(* IEC 61131-3 sources: Repository_IEMA_Test/LMC_PacDrive.device.xml.v3^/Plc Logic.plclogic.xml.v3^/Application.application.xml.v3^/TemplateFullProgrammingFramework/Examples/ExampleLeafModule/FB_ExampleLeafModule.pou.xml.v3^, 16 files *)

(* ---- Auto_Action.act.st ---- *)
__METADATA__
{
  "v3Meta": {
    "objectGuid": "52a75849-8094-4c85-bfe0-08668a2e7324",
    "objectTypeGuid": "8ac092e5-3128-4e26-9e7e-11016c6684f2",
    "embeddedObjectTypeGuids": [
      "3b83b776-fb25-43b8-99f2-3c507c9143fc"
    ],
    "properties": {},
    "subObjects": {}
  }
}

(* Start application code *)
IF(iq_stExampleLeafModuleItf.q_etState = ET_ExampleLeafModuleState.AutoWaitForStart) THEN
	IF(xAutoEnable) THEN
		IF(xStartFlag) THEN
			iq_stExampleLeafModuleItf.q_etState := ET_ExampleLeafModuleState.AutoRunning;
		END_IF
	ELSE
		xAutoActive := FALSE;
	END_IF
END_IF

IF(NOT xStartFlag AND iq_stExampleLeafModuleItf.q_etState = ET_ExampleLeafModuleState.AutoRunning) THEN
	iq_stExampleLeafModuleItf.q_etState := ET_ExampleLeafModuleState.AutoWaitForStart;
END_IF

IF(iq_stExampleLeafModuleItf.q_etState = ET_ExampleLeafModuleState.AutoRunning) THEN
	IF(xAutoEnable) THEN
		iq_stExampleLeafModuleItf.q_xValue := ifRefActualValuesPosition.RefPosition >= iq_stExampleLeafModuleItf.i_lrPosMin AND
													ifRefActualValuesPosition.RefPosition <= iq_stExampleLeafModuleItf.i_lrPosMax;
	ELSE
		iq_stExampleLeafModuleItf.q_etState := ET_ExampleLeafModuleState.AutoWaitForStart;
	END_IF
END_IF
(* End application code *)

(* ---- CancelException.meth.st ---- *)
METHOD CancelException
VAR_IN_OUT
	iq_stException	: TPL.ST_Exception;
END_VAR

TPL.FC_SetException(	i_xExceptionActive	:= FALSE,
						iq_stException		:= iq_stException,
						iq_stExceptionList	:= iq_stExceptionList,
						iq_stLogDataList	:= iq_stLogDataList,
						q_etDiag 			=> etDiagBuffer,
						q_etDiagExt 		=> etDiagExtBufferTPL,
						q_sMsg 				=> sDiagMsgBuffer);

(* ---- CheckCmd.act.st ---- *)
__METADATA__
{
  "v3Meta": {
    "objectGuid": "c3140d7a-2c8d-489a-98e5-cdbf2202bc2d",
    "objectTypeGuid": "8ac092e5-3128-4e26-9e7e-11016c6684f2",
    "embeddedObjectTypeGuids": [
      "3b83b776-fb25-43b8-99f2-3c507c9143fc"
    ],
    "properties": {},
    "subObjects": {}
  }
}

(*--------------------------------------------------------------------------------------------------*)
(* CheckCMD is checking if CMD is supported by this module *)
(*--------------------------------------------------------------------------------------------------*)
xOpModeCMD			:= FALSE;
xCheckCmdException	:= FALSE;

IF 	iq_stStandardModuleItf.iq_diCMD = ET_ExampleLeafModuleCmd.Homing OR
	iq_stStandardModuleItf.iq_diCMD = ET_ExampleLeafModuleCmd.Auto OR
	iq_stStandardModuleItf.iq_diCMD = ET_ExampleLeafModuleCmd.Stop THEN

	xOpModeCMD := TRUE;
ELSIF iq_stStandardModuleItf.iq_diCMD = ET_ExampleLeafModuleCmd.Start OR
	  iq_stStandardModuleItf.iq_diCMD = ET_ExampleLeafModuleCmd.Hold THEN
	;
ELSE
	xCheckCmdException := TRUE;
END_IF

(* ---- CmdControl_Action.act.st ---- *)
__METADATA__
{
  "v3Meta": {
    "objectGuid": "3f09c16f-6d17-42bf-986b-7819269a7b76",
    "objectTypeGuid": "8ac092e5-3128-4e26-9e7e-11016c6684f2",
    "embeddedObjectTypeGuids": [
      "3b83b776-fb25-43b8-99f2-3c507c9143fc"
    ],
    "properties": {},
    "subObjects": {}
  }
}

(* CMD execution

	algorithm:
	----------

	detect new command?
		check command?
			execute command;
		end
	end

	is command running (at least one cycle)?
		is command finished?
			signal success/unsuccessful
		end
	end
*)

xCommandAcceptedInThisCycle := FALSE;

(* Detect new command *)
IF(iq_stStandardModuleItf.i_xEnable) THEN
	IF (iq_stStandardModuleItf.iq_diCMD > 0 AND (NOT iq_stStandardModuleItf.q_xCMDActive (* In case no command is active *)
			OR iq_stStandardModuleItf.iq_diCMD <> iq_stStandardModuleItf.q_diCMDActive) (* In case a command is active *)) THEN

		xCommandRefused := FALSE; (* Flag is set by RefuseCommand() action *)

		(* Check command *)
		CheckCmd();
		IF(xCheckCmdException) THEN
			(*** Check for unknown command ***)
			stExceptionCmdUnknown.sMsg := Standard.CONCAT('Cmd unknown: ',DINT_TO_STRING(iq_stStandardModuleItf.iq_diCmd));
			ReportException(iq_stException := stExceptionCmdUnknown);
			RefuseCommand();
		ELSE
			(*** Check for impossible overwrite ***)
			IF(iq_stStandardModuleItf.q_xCMDActive AND iq_stStandardModuleItf.iq_diCMD <> ET_ExampleLeafModuleCmd.Stop) THEN (* In this module only the ET_ExampleLeafModuleCmd.Stop command can overwrite other commands *)
				stExceptionCmdImpossibleOverwrite.sMsg := PDL.FC_MultiConcat(	i_sString1 := 'Cmd impossible: ',
																				i_sString2 := FC_EtExampleLeafModuleCmdToString(i_diCmd := iq_stStandardModuleItf.iq_diCmd),
																				i_sString3 := '; Cmd active: ',
																				i_sString4 := FC_EtExampleLeafModuleCmdToString(i_diCmd := iq_stStandardModuleItf.q_diCmdActive) );
				ReportException(iq_stException := stExceptionCmdImpossibleOverwrite);
				RefuseCommand();
			ELSE
				(*** Check for impossible state ***)
				IF(NOT xOpModeCmd AND (* In this module, all OpMode commands are always possible independent of the state *)
					(iq_stExampleLeafModuleItf.q_etState = ET_ExampleLeafModuleState.NoOp (* Start and Hold are not possible in NoOp *)
					OR (iq_stExampleLeafModuleItf.q_etState = ET_ExampleLeafModuleState.HomingWaitForStart OR iq_stExampleLeafModuleItf.q_etState = ET_ExampleLeafModuleState.HomingDone) AND iq_stStandardModuleItf.iq_diCMD = ET_ExampleLeafModuleCmd.Hold) (* Hold is not supported in homing *)
					) THEN
					stExceptionCmdImpossibleState.sMsg := PDL.FC_MultiConcat(	i_sString1 := 'Cmd impossible: ',
																				i_sString2 := FC_EtExampleLeafModuleCmdToString(i_diCmd := iq_stStandardModuleItf.iq_diCmd),
																				i_sString3 := '; State: ',
																				i_sString4 := FC_EtExampleLeafModuleStateToString(i_etState := iq_stExampleLeafModuleItf.q_etState) );
					ReportException(iq_stException := stExceptionCmdImpossibleState);
					RefuseCommand();
				ELSE
					(* Check for impossible commands due to active error reactions *)
					IF	iq_stStandardModuleItf.iq_diCMD = ET_ExampleLeafModuleCmd.Start
							AND (stModuleReaction.axReaction[TPL.ET_Reaction.AsyncStop] OR
								 stModuleReaction.axReaction[TPL.ET_Reaction.SyncStopEH] OR
								 stModuleReaction.axReaction[TPL.ET_Reaction.SyncStopEL] OR
								 stModuleReaction.axReaction[TPL.ET_Reaction.StopEndOfCycle]) (* Start impossible if error reaction 4 or higher *)
						OR

						iq_stStandardModuleItf.iq_diCMD <> ET_ExampleLeafModuleCmd.Stop
							AND (stModuleReaction.axReaction[TPL.ET_Reaction.AsyncStop] OR
								 stModuleReaction.axReaction[TPL.ET_Reaction.SyncStopEH] OR
								 stModuleReaction.axReaction[TPL.ET_Reaction.SyncStopEL]) THEN (* Everything else, with exception of Stop, impossible if error reaction 3 or higher *)

						stWarningCmdImpossibleReaction.sMsg := PDL.FC_MultiConcat(	i_sString1 := 'Cmd impossible: ',
																					i_sString2 := FC_EtExampleLeafModuleCmdToString(i_diCmd := iq_stStandardModuleItf.iq_diCmd),
																					i_sString3 := '; Reaction: ',
																					i_sString4 := TPL.FC_GetStandardReactionName(iq_stReaction := stModuleReaction));
						ReportException(iq_stException := stWarningCmdImpossibleReaction);
						RefuseCommand();
					END_IF
				END_IF
			END_IF
		END_IF

		IF(NOT xCommandRefused) THEN (* Command has passed all checks, execute command *)
			IF fbLoggerPoint.etLogLevel >= APL.ET_LogLevel.UserAction THEN
				fbLoggerPoint.AddLogEntry(	i_etLogLevel	:= APL.ET_LogLevel.UserAction,
											i_etDiag		:= GD.ET_Diag.Ok,
											i_udiDiagExt	:= ET_DiagExtExampleLeafModule.Ok,
											i_sMessage		:= Standard.CONCAT(Standard.CONCAT(Standard.CONCAT('Command executing: ', FC_etExampleLeafModuleCmdToString(i_diCmd := iq_stStandardModuleItf.iq_diCmd)),' number: '),DINT_TO_STRING(iq_stStandardModuleItf.iq_diCmd)),
											q_etDiag		:= ,
											q_etDiagExt		:= );
			END_IF
			(* Accept command *)
			iq_stStandardModuleItf.q_xCMDActive := TRUE;
			iq_stStandardModuleItf.q_xCMDDone := FALSE;
			iq_stStandardModuleItf.q_diCMDActive := iq_stStandardModuleItf.iq_diCMD;

			xCommandAcceptedInThisCycle := TRUE; (* Signal for command done checks *)

			IF(xOpModeCMD) THEN
				DisableAllJobs();

				CASE iq_stStandardModuleItf.iq_diCMD OF
					ET_ExampleLeafModuleCmd.Stop:
						;	(* Do nothing, disabled OpMode flags automatically lead to NoOp *)

					ET_ExampleLeafModuleCmd.Homing:
						xHomingEnable := TRUE;

					ET_ExampleLeafModuleCmd.Auto:
						xAutoEnable := TRUE;
				END_CASE
			ELSE
				(* Action commands *)
				CASE iq_stStandardModuleItf.iq_diCMD OF
					ET_ExampleLeafModuleCmd.Start:
						xStartFlag := TRUE;

					ET_ExampleLeafModuleCmd.Hold:
						xStartFlag := FALSE;
				END_CASE
			END_IF
		END_IF (* New command? *)
	END_IF

(********************************************* Check successful and unsucessful of given commands ****************************************)

	(* Check if active command is done or is stopped by an error *)
	IF(NOT xCommandAcceptedInThisCycle) THEN (* Don't execute these checks if we accepted a new command in this cycle
		to ensure that execution of every command requires a minimum of 2 cycles *)

		IF(iq_stStandardModuleItf.q_xCMDActive) THEN
			CASE iq_stStandardModuleItf.iq_diCmd OF
				ET_ExampleLeafModuleCmd.Homing:
					(* Successful *)
					IF(xHomingActive) THEN
						SignalSuccessfulExecution();
					END_IF
					(* Unsucessful *)
					IF (stModuleReaction.axReaction[TPL.ET_Reaction.AsyncStop] OR
						stModuleReaction.axReaction[TPL.ET_Reaction.SyncStopEL] OR
						stModuleReaction.axReaction[TPL.ET_Reaction.SyncStopEH]) THEN

						SignalUnsuccessfulExecution();
					END_IF

				ET_ExampleLeafModuleCmd.Auto:
					(* Successful *)
					IF(xAutoActive) THEN
						SignalSuccessfulExecution();
					END_IF
					(* Unsucessful *)
					IF (stModuleReaction.axReaction[TPL.ET_Reaction.AsyncStop] OR
						stModuleReaction.axReaction[TPL.ET_Reaction.SyncStopEL] OR
						stModuleReaction.axReaction[TPL.ET_Reaction.SyncStopEH]) THEN

						SignalUnsuccessfulExecution();
					END_IF

				ET_ExampleLeafModuleCmd.Stop:
					(* Successful *)
					IF(iq_stExampleLeafModuleItf.q_etState = ET_ExampleLeafModuleState.NoOp) THEN
						SignalSuccessfulExecution();
					END_IF

				ET_ExampleLeafModuleCmd.Start:
					IF(iq_stExampleLeafModuleItf.q_etState = ET_ExampleLeafModuleState.HomingDone) THEN
						xStartFlag := FALSE;
					END_IF
					(* Successful *)
					IF(iq_stExampleLeafModuleItf.q_etState = ET_ExampleLeafModuleState.HomingDone AND NOT xHomingException
						OR iq_stExampleLeafModuleItf.q_etState = ET_ExampleLeafModuleState.AutoRunning) THEN
						SignalSuccessfulExecution();
					END_IF
					(* Unsucessful *)
					IF (stModuleReaction.axReaction[TPL.ET_Reaction.AsyncStop] OR
						stModuleReaction.axReaction[TPL.ET_Reaction.SyncStopEL] OR
						stModuleReaction.axReaction[TPL.ET_Reaction.SyncStopEH] OR
						stModuleReaction.axReaction[TPL.ET_Reaction.StopEndOfCycle]  OR
						iq_stExampleLeafModuleItf.q_etState = ET_ExampleLeafModuleState.HomingDone AND xHomingException) THEN

						SignalUnsuccessfulExecution();
					END_IF

				ET_ExampleLeafModuleCmd.Hold:
					(* Successful *)
					IF(iq_stExampleLeafModuleItf.q_etState = ET_ExampleLeafModuleState.AutoWaitForStart) THEN
						SignalSuccessfulExecution();
					END_IF
					(* Unsucessful *)
					IF (stModuleReaction.axReaction[TPL.ET_Reaction.AsyncStop] OR
						stModuleReaction.axReaction[TPL.ET_Reaction.SyncStopEL] OR
						stModuleReaction.axReaction[TPL.ET_Reaction.SyncStopEH]) THEN

						SignalUnsuccessfulExecution();
					END_IF
			END_CASE
		END_IF
	END_IF
ELSE
	(* Module is going to be disabled *)
	iq_stStandardModuleItf.q_xReady := FALSE;
	xEnableFlag := FALSE;

	DisableAllJobs();

	xStartFlag := FALSE;

	IF(iq_stStandardModuleItf.q_xCmdActive) THEN (* If a command is currently active, cancel its execution *)
		SignalUnsuccessfulExecution();
	ELSE
		InactiveCmdExecution(); (* Command processing as if we were disabled *)
	END_IF
END_IF

(* ---- DiagQuit.act.st ---- *)
__METADATA__
{
  "v3Meta": {
    "objectGuid": "69ccc72d-2ac0-4551-ad4e-f7cbec51c7c2",
    "objectTypeGuid": "8ac092e5-3128-4e26-9e7e-11016c6684f2",
    "embeddedObjectTypeGuids": [
      "3b83b776-fb25-43b8-99f2-3c507c9143fc"
    ],
    "properties": {},
    "subObjects": {}
  }
}

IF(iq_stStandardModuleItf.i_xDiagQuit AND NOT xDiagQuitFlag) THEN
	(* Rising edge of error quit *)
	xDiagQuitFlag := TRUE;
	xNotAbleToSetException := FALSE;

	FOR udii := 1 TO TPL.ET_Reaction.MainsContactorOff DO
		stLocalReaction.axReaction[udii] := FALSE;
	END_FOR

	iq_stStandardModuleItf.q_etDiag := GD.ET_Diag.Ok;

	IF(iq_stStandardModuleItf.iq_diCMD < 0) THEN
		iq_stStandardModuleItf.iq_diCMD := 0;
	END_IF
	IF fbLoggerPoint.etLogLevel >= APL.ET_LogLevel.UserAction THEN
		fbLoggerPoint.AddLogEntry(	i_etLogLevel	:= APL.ET_LogLevel.UserAction,
									i_etDiag		:= GD.ET_Diag.Ok,
									i_udiDiagExt	:= ET_DiagExtExampleLeafModule.Ok,
									i_sMessage		:= 'Diag Quit',
									q_etDiag		:= ,
									q_etDiagExt		:= );
	END_IF
ELSIF(NOT iq_stStandardModuleItf.i_xDiagQuit AND xDiagQuitFlag) THEN
	xDiagQuitFlag := FALSE;
END_IF

(* ---- ExceptionHandler_Action.act.st ---- *)
__METADATA__
{
  "v3Meta": {
    "objectGuid": "988a9a77-f250-4378-92cf-5dc7496f5b9c",
    "objectTypeGuid": "8ac092e5-3128-4e26-9e7e-11016c6684f2",
    "embeddedObjectTypeGuids": [
      "3b83b776-fb25-43b8-99f2-3c507c9143fc"
    ],
    "properties": {},
    "subObjects": {}
  }
}

(* -----------------------------------------------------------------------------------------------*)
(* Check Axis Errors *)
(* -----------------------------------------------------------------------------------------------*)
	IF (iq_stExampleLeafModuleItf.i_ifDrive.DiagClass > 3) THEN
		stExceptionDriveFatal.sMsg := PDL.FC_MultiConcat(	i_sString1 := 'DiagCode: ',
															i_sString2 := DINT_TO_STRING(iq_stExampleLeafModuleItf.i_ifDrive.DiagCode),
															i_sString3 := ' Msg: ',
															i_sString4 := iq_stExampleLeafModuleItf.i_ifDrive.DiagMsg);

		ReportException(iq_stException := stExceptionDriveFatal);

	ELSIF (iq_stExampleLeafModuleItf.i_ifDrive.DiagClass = 3) THEN
		stExcepitonDrive.sMsg := PDL.FC_MultiConcat(	i_sString1 := 'DiagCode: ',
														i_sString2 := DINT_TO_STRING(iq_stExampleLeafModuleItf.i_ifDrive.DiagCode),
														i_sString3 := ' Msg: ',
														i_sString4 := iq_stExampleLeafModuleItf.i_ifDrive.DiagMsg);

		ReportException(iq_stException := stExcepitonDrive);

	ELSIF (iq_stExampleLeafModuleItf.i_ifDrive.DiagClass > 0)  AND (iq_stExampleLeafModuleItf.i_ifDrive.DiagClass < 3) THEN
		stWarningDrive.sMsg := PDL.FC_MultiConcat(	i_sString1 := 'DiagCode: ',
													i_sString2 := DINT_TO_STRING(iq_stExampleLeafModuleItf.i_ifDrive.DiagCode),
													i_sString3 := ' Msg: ',
													i_sString4 := iq_stExampleLeafModuleItf.i_ifDrive.DiagMsg);

		ReportException(iq_stException := stWarningDrive);
	END_IF

(* -----------------------------------------------------------------------------------------------*)
(* Check StopModi *)
(* -----------------------------------------------------------------------------------------------*)
IF (NOT iq_stStandardModuleItf.i_xEnable OR
	stModuleReaction.axReaction[TPL.ET_Reaction.AsyncStop] OR
	stModuleReaction.axReaction[TPL.ET_Reaction.SyncStopEL] OR
	stModuleReaction.axReaction[TPL.ET_Reaction.SyncStopEH]) THEN

	xAutoEnable := FALSE;
	xHomingEnable := FALSE;
END_IF
IF (NOT iq_stStandardModuleItf.i_xEnable OR
	stModuleReaction.axReaction[TPL.ET_Reaction.AsyncStop] OR
	stModuleReaction.axReaction[TPL.ET_Reaction.SyncStopEL] OR
	stModuleReaction.axReaction[TPL.ET_Reaction.SyncStopEH] OR
	stModuleReaction.axReaction[TPL.ET_Reaction.StopEndOfCycle] ) THEN

	xStartFlag := FALSE;
END_IF

(* ---- Homing_Action.act.st ---- *)
__METADATA__
{
  "v3Meta": {
    "objectGuid": "1a034643-a971-4ebb-a9e0-a35821b4c802",
    "objectTypeGuid": "8ac092e5-3128-4e26-9e7e-11016c6684f2",
    "embeddedObjectTypeGuids": [
      "3b83b776-fb25-43b8-99f2-3c507c9143fc"
    ],
    "properties": {},
    "subObjects": {}
  }
}

(* Start application code *)
IF(xStartFlag AND (iq_stExampleLeafModuleItf.q_etState = ET_ExampleLeafModuleState.HomingWaitForStart OR iq_stExampleLeafModuleItf.q_etState = ET_ExampleLeafModuleState.HomingDone)) THEN
	xHomingException := FALSE;
	iq_stExampleLeafModuleItf.q_etState := ET_ExampleLeafModuleState.HomingExecuting;
END_IF

IF(iq_stExampleLeafModuleItf.q_etState = ET_ExampleLeafModuleState.HomingExecuting) THEN
	(* Emulating an action in the process that takes some time *)
	udiDoSomethingCounter := udiDoSomethingCounter + 1;
	IF(udiDoSomethingCounter > c_udiDoSomeThingLevel) THEN
		(* Homing done *)
		iq_stExampleLeafModuleItf.q_xValue := TRUE;

		(* Sometimes creates an error *)
		IF(iq_stExampleLeafModuleItf.i_xEnableRandomExceptionTrigger) THEN
			IF(xRandomExceptionTrigger) THEN
				xHomingException := TRUE;
			END_IF
			xRandomExceptionTrigger := NOT xRandomExceptionTrigger;
		END_IF

		iq_stExampleLeafModuleItf.q_etState := ET_ExampleLeafModuleState.HomingDone;
	END_IF
END_IF

IF xHomingException THEN
	ReportException(iq_stException := stExceptionHoming);
ELSE
	CancelException(iq_stException := stExceptionHoming);
END_IF

IF(iq_stExampleLeafModuleItf.q_etState <> ET_ExampleLeafModuleState.HomingExecuting) THEN
	(* If homing is not running, allow exit of homing by xHomingEnable = FALSE *)
	IF(NOT xHomingEnable) THEN
		xHomingActive := FALSE;
	END_IF
END_IF
(* End application code *)

(* ---- InactiveCmdExecution.act.st ---- *)
__METADATA__
{
  "v3Meta": {
    "objectGuid": "2d98f9c2-2241-4178-a153-8519baf7c94c",
    "objectTypeGuid": "8ac092e5-3128-4e26-9e7e-11016c6684f2",
    "embeddedObjectTypeGuids": [
      "3b83b776-fb25-43b8-99f2-3c507c9143fc"
    ],
    "properties": {},
    "subObjects": {}
  }
}

(* Command execution if module is not active (q_xActive = FALSE) or currently deactivating (i_xEnable = FALSE, q_xActive is still TRUE) *)
IF iq_stStandardModuleItf.iq_diCmd <> 0 THEN
	IF(NOT iq_stStandardModuleItf.i_xEnable) THEN
		iq_stStandardModuleItf.iq_diCmd := 0; (* All commands are signaled executed if module is disabled *)
(*ELSE*)
	ELSIF(iq_stStandardModuleItf.iq_diCmd > 0) THEN (* New command *)
		(* Command execution during enable but module is not ready for commands yet ==> error *)
		//xExceptionCmdImpossibleState := TRUE;

		stExceptionCmdImpossibleState.sMsg := PDL.FC_MultiConcat(	i_sString1 := 'Cmd impossible: ',
																	i_sString2 := FC_EtExampleLeafModuleCmdToString(i_diCmd := ABS(iq_stStandardModuleItf.iq_diCmd)),
																	i_sString3 := '; State: ',
																	i_sString4 := FC_EtExampleLeafModuleStateToString(i_etState := iq_stExampleLeafModuleItf.q_etState));
		ReportException(iq_stException := stExceptionCmdImpossibleState);
		iq_stStandardModuleItf.iq_diCmd:= - ABS(iq_stStandardModuleItf.iq_diCmd);
	END_IF
END_IF
iq_stStandardModuleItf.q_xCmdActive := FALSE;
iq_stStandardModuleItf.q_xCmdDone := FALSE;
iq_stStandardModuleItf.q_diCmdActive := 0;

(* ---- Init_Action.act.st ---- *)
__METADATA__
{
  "v3Meta": {
    "objectGuid": "be2905dd-e781-480e-b168-a410b5083870",
    "objectTypeGuid": "8ac092e5-3128-4e26-9e7e-11016c6684f2",
    "embeddedObjectTypeGuids": [
      "3b83b776-fb25-43b8-99f2-3c507c9143fc"
    ],
    "properties": {},
    "subObjects": {}
  }
}

iq_stStandardModuleItf.q_xActive			:= FALSE;
iq_stStandardModuleItf.q_xReady				:= FALSE;

iq_stStandardModuleItf.q_etDiag				:= GD.ET_Diag.Ok;
iq_stStandardModuleItf.q_udiDiagExt			:= ET_DiagExtExampleLeafModule.Disabled;
iq_stStandardModuleItf.q_sDiagExt			:= FC_EtDiagExtExampleLeafModuleToString(i_etDiagExt := iq_stStandardModuleItf.q_udiDiagExt);
iq_stStandardModuleItf.q_sMsg				:= '';

iq_stStandardModuleItf.q_dwModuleType		:= ET_ModuleType.ExampleLeafModule;
iq_stStandardModuleItf.q_sModuleTypeName	:= 'ExampleLeafModule';
iq_stStandardModuleItf.q_udiModuleVersion	:= 1;

iq_stExampleLeafModuleItf.q_etState	:= ET_ExampleLeafModuleState.Disabled;

THIS^.DiagQuit();
THIS^.InactiveCmdExecution();

udiMyResultSource := ET_ExceptionSource.ExampleLeafModule; (* Has to be coded this way to get around compiler restrictions*)

(* detect invalid configurations and avoid array index out of range error *)
IF(iq_stStandardModuleItf.iq_stExt.udiReactionOffset + TPL. ET_Reaction.MainsContactorOff > TPL.Gc_udiMaxNumberOfReactions) OR xExceptionReactionOutsideRange THEN (* module uses error reactions 1 to 5 *)
	xExceptionReactionOutsideRange := TRUE; (* create unquittable error *)

	(* create exception *)
	stExceptionInit.etDiag					:= GD.ET_Diag.InputParameterInvalid;
	stExceptionInit.udiDiagExt				:= ET_DiagExtExampleLeafModule.ReactionOffsetRange;
	stExceptionInit.sMsg					:= Standard.CONCAT('Value: ', UDINT_TO_STRING(iq_stStandardModuleItf.iq_stExt.udiReactionOffset));
	stExceptionInit.udiModuleId				:= iq_stStandardModuleItf.i_udiModuleId;
	stExceptionInit.sModuleName				:= iq_stStandardModuleItf.i_sModuleName;
	stExceptionInit.etSource				:= udiMyResultSource;
	stExceptionInit.timDelayTime			:= T#0MS;
	stExceptionInit.wHmiAttributes			:= 0;
	stExceptionInit.xAutoQuit				:= FALSE;
	stExceptionInit.stReaction.axReaction[TPL.ET_Reaction.AsyncStop]	:= TRUE; (* without offset on purpose *)

	iq_stStandardModuleItf.iq_stExt.udiReactionOffset := 0;

	ReportException(iq_stException := stExceptionInit);
ELSIF (iq_stStandardModuleItf.i_xEnable) THEN
	stReaction1 := stEmptyReaction;
	stReaction1.axReaction[iq_stStandardModuleItf.iq_stExt.udiReactionOffset + TPL.ET_Reaction.AsyncStop] := TRUE;
	stReaction2 := stEmptyReaction;
	stReaction2.axReaction[iq_stStandardModuleItf.iq_stExt.udiReactionOffset + TPL.ET_Reaction.SyncStopEL] := TRUE;
	stReaction3 := stEmptyReaction;
	stReaction3.axReaction[iq_stStandardModuleItf.iq_stExt.udiReactionOffset + TPL.ET_Reaction.SyncStopEH] := TRUE;
	stReaction4 := stEmptyReaction;
	stReaction4.axReaction[iq_stStandardModuleItf.iq_stExt.udiReactionOffset + TPL.ET_Reaction.StopEndOfCycle] := TRUE;

	(* Initialization of exception structures *)
	stExceptionCmdUnknown.etDiag						:= GD.ET_Diag.ExecutionAborted;
	stExceptionCmdUnknown.udiDiagExt					:= ET_DiagExtExampleLeafModule.CmdUnknown;
	stExceptionCmdUnknown.sMsg							:= 'Command unknown'; (* Replaced on usage *)
	stExceptionCmdUnknown.udiModuleId					:= iq_stStandardModuleItf.i_udiModuleId;
	stExceptionCmdUnknown.sModuleName					:= iq_stStandardModuleItf.i_sModuleName;
	stExceptionCmdUnknown.etSource						:= udiMyResultSource;
	stExceptionCmdUnknown.timDelayTime					:= T#0MS;
	stExceptionCmdUnknown.wHmiAttributes				:= 0;
	stExceptionCmdUnknown.xAutoQuit						:= FALSE;
	stExceptionCmdUnknown.stReaction					:= stReaction1;

	stExceptionCmdImpossibleOverwrite.etDiag			:= GD.ET_Diag.ExecutionAborted;
	stExceptionCmdImpossibleOverwrite.udiDiagExt		:= ET_DiagExtExampleLeafModule.CmdImpossibleOverwrite;
	stExceptionCmdImpossibleOverwrite.sMsg				:= 'Impossible command overwrite'; (* Replaced on usage *)
	stExceptionCmdImpossibleOverwrite.udiModuleId		:= iq_stStandardModuleItf.i_udiModuleId;
	stExceptionCmdImpossibleOverwrite.sModuleName		:= iq_stStandardModuleItf.i_sModuleName;
	stExceptionCmdImpossibleOverwrite.etSource			:= udiMyResultSource;
	stExceptionCmdImpossibleOverwrite.timDelayTime		:= T#0MS;
	stExceptionCmdImpossibleOverwrite.wHmiAttributes	:= 0;
	stExceptionCmdImpossibleOverwrite.xAutoQuit			:= FALSE;
	stExceptionCmdImpossibleOverwrite.stReaction		:= stReaction1;

	stExceptionCmdImpossibleState.etDiag				:= GD.ET_Diag.ExecutionAborted;
	stExceptionCmdImpossibleState.udiDiagExt			:= ET_DiagExtExampleLeafModule.CmdImpossibleState;
	stExceptionCmdImpossibleState.sMsg					:= 'Impossible command for state'; (* Replaced on usage *)
	stExceptionCmdImpossibleState.udiModuleId			:= iq_stStandardModuleItf.i_udiModuleId;
	stExceptionCmdImpossibleState.sModuleName			:= iq_stStandardModuleItf.i_sModuleName;
	stExceptionCmdImpossibleState.etSource				:= udiMyResultSource;
	stExceptionCmdImpossibleState.timDelayTime			:= T#0MS;
	stExceptionCmdImpossibleState.wHmiAttributes		:= 0;
	stExceptionCmdImpossibleState.xAutoQuit				:= FALSE;
	stExceptionCmdImpossibleState.stReaction			:= stReaction1;

	stWarningCmdImpossibleReaction.etDiag				:= GD.ET_Diag.ExecutionAborted;
	stWarningCmdImpossibleReaction.udiDiagExt			:= ET_DiagExtExampleLeafModule.CmdImpossibleReaction;
	stWarningCmdImpossibleReaction.sMsg					:= 'Impossible command on reaction'; (* Replaced on usage *)
	stWarningCmdImpossibleReaction.udiModuleId			:= iq_stStandardModuleItf.i_udiModuleId;
	stWarningCmdImpossibleReaction.sModuleName			:= iq_stStandardModuleItf.i_sModuleName;
	stWarningCmdImpossibleReaction.etSource				:= udiMyResultSource;
	stWarningCmdImpossibleReaction.timDelayTime			:= T#0MS;
	stWarningCmdImpossibleReaction.wHmiAttributes		:= 0;
	stWarningCmdImpossibleReaction.xAutoQuit			:= FALSE;

	stExceptionModuleReaction1.etDiag					:= GD.ET_Diag.InputParameterInvalid;(* Replaced on usage *)
	stExceptionModuleReaction1.udiDiagExt				:= ET_DiagExtExampleLeafModule.Ok;(* Replaced on usage *)
	stExceptionModuleReaction1.sMsg						:= '';(* Replaced on usage *)
	stExceptionModuleReaction1.udiModuleId				:= iq_stStandardModuleItf.i_udiModuleId;
	stExceptionModuleReaction1.sModuleName				:= iq_stStandardModuleItf.i_sModuleName;
	stExceptionModuleReaction1.etSource					:= udiMyResultSource;
	stExceptionModuleReaction1.timDelayTime				:= T#0MS;
	stExceptionModuleReaction1.wHmiAttributes			:= 0;
	stExceptionModuleReaction1.xAutoQuit				:= FALSE;
	stExceptionModuleReaction1.stReaction				:= stReaction1;

	stExceptionModuleReaction2.etDiag					:= GD.ET_Diag.InputParameterInvalid;(* Replaced on usage *)
	stExceptionModuleReaction2.udiDiagExt				:= ET_DiagExtExampleLeafModule.Ok;(* Replaced on usage *)
	stExceptionModuleReaction2.sMsg						:= '';(* Replaced on usage *)
	stExceptionModuleReaction2.udiModuleId				:= iq_stStandardModuleItf.i_udiModuleId;
	stExceptionModuleReaction2.sModuleName				:= iq_stStandardModuleItf.i_sModuleName;
	stExceptionModuleReaction2.etSource					:= udiMyResultSource;
	stExceptionModuleReaction2.timDelayTime				:= T#0MS;
	stExceptionModuleReaction2.wHmiAttributes			:= 0;
	stExceptionModuleReaction2.xAutoQuit				:= FALSE;
	stExceptionModuleReaction2.stReaction				:= stReaction2;

	stExceptionModuleReaction3.etDiag					:= GD.ET_Diag.InputParameterInvalid;(* Replaced on usage *)
	stExceptionModuleReaction3.udiDiagExt				:= ET_DiagExtExampleLeafModule.Ok;(* Replaced on usage *)
	stExceptionModuleReaction3.sMsg						:= '';(* Replaced on usage *)
	stExceptionModuleReaction3.udiModuleId				:= iq_stStandardModuleItf.i_udiModuleId;
	stExceptionModuleReaction3.sModuleName				:= iq_stStandardModuleItf.i_sModuleName;
	stExceptionModuleReaction3.etSource					:= udiMyResultSource;
	stExceptionModuleReaction3.timDelayTime				:= T#0MS;
	stExceptionModuleReaction3.wHmiAttributes			:= 0;
	stExceptionModuleReaction3.xAutoQuit				:= FALSE;
	stExceptionModuleReaction3.stReaction				:= stReaction3;

	stExceptionModuleReaction4.etDiag					:= GD.ET_Diag.InputParameterInvalid;(* Replaced on usage *)
	stExceptionModuleReaction4.udiDiagExt				:= ET_DiagExtExampleLeafModule.Ok;(* Replaced on usage *)
	stExceptionModuleReaction4.sMsg						:= '';(* Replaced on usage *)
	stExceptionModuleReaction4.udiModuleId				:= iq_stStandardModuleItf.i_udiModuleId;
	stExceptionModuleReaction4.sModuleName				:= iq_stStandardModuleItf.i_sModuleName;
	stExceptionModuleReaction4.etSource					:= udiMyResultSource;
	stExceptionModuleReaction4.timDelayTime				:= T#0MS;
	stExceptionModuleReaction4.wHmiAttributes			:= 0;
	stExceptionModuleReaction4.xAutoQuit				:= FALSE;
	stExceptionModuleReaction4.stReaction				:= stReaction4;

	stExceptionDriveFatal.etDiag						:= GD.ET_Diag.DriveConditionInvalid;
	stExceptionDriveFatal.udiDiagExt					:= ET_DiagExtExampleLeafModule.DriveFatalException;
	stExceptionDriveFatal.sMsg							:= 'Drive diag'; (* Replaced on usage *)
	stExceptionDriveFatal.udiModuleId					:= iq_stStandardModuleItf.i_udiModuleId;
	stExceptionDriveFatal.sModuleName					:= iq_stStandardModuleItf.i_sModuleName;
	stExceptionDriveFatal.etSource						:= udiMyResultSource;
	stExceptionDriveFatal.timDelayTime					:= T#0MS;
	stExceptionDriveFatal.wHmiAttributes				:= 0;
	stExceptionDriveFatal.xAutoQuit						:= FALSE;
	stExceptionDriveFatal.stReaction					:= stReaction1;

	stExcepitonDrive.etDiag								:= GD.ET_Diag.DriveConditionInvalid;
	stExcepitonDrive.udiDiagExt							:= ET_DiagExtExampleLeafModule.DriveException;
	stExcepitonDrive.sMsg								:= 'Drive diag'; (* Replaced on usage *)
	stExcepitonDrive.udiModuleId						:= iq_stStandardModuleItf.i_udiModuleId;
	stExcepitonDrive.sModuleName						:= iq_stStandardModuleItf.i_sModuleName;
	stExcepitonDrive.etSource							:= udiMyResultSource;
	stExcepitonDrive.timDelayTime						:= T#0MS;
	stExcepitonDrive.wHmiAttributes						:= 0;
	stExcepitonDrive.xAutoQuit							:= FALSE;
	stExcepitonDrive.stReaction							:= stReaction2;

	stWarningDrive.etDiag								:= GD.ET_Diag.DriveConditionInvalid;
	stWarningDrive.udiDiagExt							:= ET_DiagExtExampleLeafModule.DriveWarning;
	stWarningDrive.sMsg									:= 'Drive warning'; (* Replaced on usage *)
	stWarningDrive.udiModuleId							:= iq_stStandardModuleItf.i_udiModuleId;
	stWarningDrive.sModuleName							:= iq_stStandardModuleItf.i_sModuleName;
	stWarningDrive.etSource								:= udiMyResultSource;
	stWarningDrive.timDelayTime							:= T#0MS;
	stWarningDrive.wHmiAttributes						:= 0;
	stWarningDrive.xAutoQuit							:= FALSE;
	stWarningDrive.stReaction							:= stReaction4;

	stExceptionInit.etDiag								:= GD.ET_Diag.InputParameterInvalid; (* Replaced on usage *)
	stExceptionInit.udiDiagExt							:= ET_DiagExtExampleLeafModule.Ok; (* Replaced on usage *)
	stExceptionInit.sMsg								:= ''; (* Replaced on usage *)
	stExceptionInit.udiModuleId							:= iq_stStandardModuleItf.i_udiModuleId;
	stExceptionInit.sModuleName							:= iq_stStandardModuleItf.i_sModuleName;
	stExceptionInit.etSource							:= udiMyResultSource;
	stExceptionInit.timDelayTime						:= T#0MS;
	stExceptionInit.wHmiAttributes						:= 0;
	stExceptionInit.xAutoQuit							:= FALSE;
	stExceptionInit.stReaction							:= stReaction1;

	stExceptionHoming.etDiag							:= GD.ET_Diag.HomingFailed;
	stExceptionHoming.udiDiagExt						:= ET_DiagExtExampleLeafModule.RandomException;
	stExceptionHoming.sMsg								:= '';
	stExceptionHoming.udiModuleId						:= iq_stStandardModuleItf.i_udiModuleId;
	stExceptionHoming.sModuleName						:= iq_stStandardModuleItf.i_sModuleName;
	stExceptionHoming.etSource							:= udiMyResultSource;
	stExceptionHoming.timDelayTime						:= T#0MS;
	stExceptionHoming.wHmiAttributes					:= 0;
	stExceptionHoming.xAutoQuit							:= FALSE;
	stExceptionHoming.stReaction						:= stReaction4;

	IF (iq_stExampleLeafModuleItf.i_ifDrive = 0) THEN
		stExceptionModuleReaction1.etDiag		:= GD.ET_Diag.InputParameterInvalid;
		stExceptionModuleReaction1.udiDiagExt	:= ET_DiagExtExampleLeafModule.DriveInvalid;
		stExceptionModuleReaction1.sMsg			:= 'No drive given';

		ReportException(iq_stException := stExceptionModuleReaction1);
	ELSE
		xEnableFlag := TRUE;
		iq_stStandardModuleItf.q_xActive := TRUE;

		FOR udii := 1 TO TPL.Gc_udiMaxNumberOfReactions DO
			stLocalReaction.axReaction[udii] := FALSE;
		END_FOR

		THIS^.SetInterfaces();

		xInitHomingDone := FALSE;

		iq_stExampleLeafModuleItf.q_etState := ET_ExampleLeafModuleState.Initializing;

		iq_stStandardModuleItf.q_etDiag		:= GD.ET_Diag.Ok;
		iq_stStandardModuleItf.q_udiDiagExt	:= ET_DiagExtExampleLeafModule.Initializing;
		iq_stStandardModuleItf.q_sDiagExt	:= FC_EtDiagExtExampleLeafModuleToString(ET_DiagExtExampleLeafModule.Initializing);
		iq_stStandardModuleItf.q_sMsg		:= '';

		IF fbLoggerPoint.etLogLevel >= APL.ET_LogLevel.UserAction THEN
			fbLoggerPoint.AddLogEntry(	i_etLogLevel	:= APL.ET_LogLevel.UserAction,
										i_etDiag		:= GD.ET_Diag.Ok,
										i_udiDiagExt	:= ET_DiagExtExampleLeafModule.Ok,
										i_sMessage		:= 'enabeling Module',
										q_etDiag		:= ,
										q_etDiagExt		:= );
		END_IF
	END_IF

END_IF

THIS^.SetOutputs();

(* ---- InitHoming_Action.act.st ---- *)
__METADATA__
{
  "v3Meta": {
    "objectGuid": "522d2040-ce61-42de-b75b-9fa026d7e50e",
    "objectTypeGuid": "8ac092e5-3128-4e26-9e7e-11016c6684f2",
    "embeddedObjectTypeGuids": [
      "3b83b776-fb25-43b8-99f2-3c507c9143fc"
    ],
    "properties": {},
    "subObjects": {}
  }
}

DiagQuit();
InactiveCmdExecution();

(* Emulating an initialization that takes some time *)
udiDoSomethingCounter := udiDoSomethingCounter + 1;
IF(iq_stExampleLeafModuleItf.i_xInitHoming) THEN
	xInitHomingDone := FALSE;
	iq_stExampleLeafModuleItf.q_xValue := TRUE;
	IF(udiDoSomethingCounter > c_udiDoSomeThingLevel) THEN
		(* Initial homing done *)
		xInitHomingDone := TRUE;
		iq_stExampleLeafModuleItf.q_xValue := TRUE;
		IF fbLoggerPoint.etLogLevel >= APL.ET_LogLevel.StatusMessage THEN
			fbLoggerPoint.AddLogEntry(	i_etLogLevel	:= APL.ET_LogLevel.StatusMessage,
										i_etDiag		:= GD.ET_Diag.Ok,
										i_udiDiagExt	:= ET_DiagExtExampleLeafModule.Ok,
										i_sMessage		:= 'InitHoming done',
										q_etDiag		:= ,
										q_etDiagExt		:= );
		END_IF
	END_IF
ELSE
	xInitHomingDone := TRUE;
END_IF

THIS^.SetOutputs();

(* ---- RegisterLoggerPoint.meth.st ---- *)
METHOD PUBLIC RegisterLoggerPoint
VAR_INPUT
	i_ifParent		: APL.IF_LoggerPoint;
	i_sName			: STRING[80];
END_VAR
VAR_OUTPUT
	q_etDiag		: GD.ET_Diag := GD.ET_Diag.Ok;
	q_etDiagExt		: ET_DiagExtExampleLeafModule := ET_DiagExtExampleLeafModule.Ok;
	q_sMsg			: STRING[80] := '';
END_VAR
VAR
	etDiagBuffer		: GD.ET_Diag;
	etDiagExtBufferAPL	: APL.ET_DiagExt;
END_VAR

THIS^.fbLoggerPoint.RegisterLoggerPoint(	i_ifParent		:= i_ifParent,
											i_sName			:= i_sName,
											i_sType			:= 'FB_ExampleLeafModule',
											i_sSource		:= 'Project',
											q_etDiag		=> etDiagBuffer,
											q_etDiagExt		=> etDiagExtBufferAPL);
IF (etDiagBuffer <> GD.ET_Diag.Ok) THEN
	CASE etDiagExtBufferAPL OF
		APL.ET_DiagExt.ParentInvalid:
			q_etDiag := GD.ET_Diag.InputParameterInvalid;
			q_etDiagExt := ET_DiagExtExampleLeafModule.ParentInvalid;

		APL.ET_DiagExt.ParentNotRegistered:
			q_etDiag := GD.ET_Diag.InputParameterInvalid;
			q_etDiagExt := ET_DiagExtExampleLeafModule.ParentNotRegistered;

		APL.ET_DiagExt.MaxNumberOfLoggerPointsExeeded:
			q_etDiag := GD.ET_Diag.InputParameterInvalid;
			q_etDiagExt := ET_DiagExtExampleLeafModule.MaxNumberOfLoggerPointsExeeded;

	ELSE
		q_etDiag := GD.ET_Diag.UnexpectedProgramBehavior;
		q_etdiagExt := ET_DiagExtExampleLeafModule.UnexpectedDiagExt;
		q_sMsg := Standard.CONCAT('RegisterLoggerPoint: ', APL.FC_EtDiagExtToString(i_etDiagExt := etDiagExtBufferAPL));
	END_CASE
END_IF

(* ---- ReportException.meth.st ---- *)
METHOD ReportException
VAR_IN_OUT
	iq_stException	: TPL.ST_Exception;
END_VAR
VAR CONSTANT
	c_diMaxReaction	: DINT := 4;
END_VAR

IF (fbLoggerPoint.etLogLevel >= APL.ET_LogLevel.CriticalException) AND (iq_stException.etDiag = GD.ET_Diag.UnexpectedProgramBehavior) THEN
	IF NOT TPL.FC_CheckExceptionIsInList( iq_stException := iq_stException, iq_stExceptionList := THIS^.iq_stExceptionList) THEN
		fbLoggerPoint.AddLogEntry(	i_etLogLevel	:= APL.ET_LogLevel.CriticalException,
									i_etDiag		:= GD.ET_Diag.Ok,
									i_udiDiagExt	:= ET_DiagExtExampleLeafModule.Ok,
									i_sMessage		:= Standard.CONCAT(Standard.CONCAT(Standard.CONCAT(Standard.CONCAT(Standard.CONCAT(Standard.CONCAT('Exception ET_Diag: ',GD.FC_EtDiagToString(i_etDiag := iq_stException.etDiag)),' ET_DiagExt: '),FC_EtDiagExtToString(i_etDiagExt := iq_stException.udiDiagExt)),' sMsg: '),iq_stException.sMsg),TPL.FC_GetStandardReactionName(iq_stReaction := iq_stException.stReaction)),
									q_etDiag		:= ,
									q_etDiagExt		:= );
	END_IF
ELSIF (fbLoggerPoint.etLogLevel >= APL.ET_LogLevel.Exception) THEN
	IF NOT TPL.FC_CheckExceptionIsInList( iq_stException := iq_stException, iq_stExceptionList := THIS^.iq_stExceptionList) THEN
		fbLoggerPoint.AddLogEntry(	i_etLogLevel	:= APL.ET_LogLevel.Exception,
									i_etDiag		:= GD.ET_Diag.Ok,
									i_udiDiagExt	:= ET_DiagExtExampleLeafModule.Ok,
									i_sMessage		:= Standard.CONCAT(Standard.CONCAT(Standard.CONCAT(Standard.CONCAT(Standard.CONCAT(Standard.CONCAT('Exception ET_Diag: ',GD.FC_EtDiagToString(i_etDiag := iq_stException.etDiag)),' ET_DiagExt: '),FC_EtDiagExtToString(i_etDiagExt := iq_stException.udiDiagExt)),' sMsg: '),iq_stException.sMsg),TPL.FC_GetStandardReactionName(iq_stReaction := iq_stException.stReaction)),
									q_etDiag		:= ,
									q_etDiagExt		:= );
	END_IF
END_IF

iq_stException.sDiagExt := FC_EtDiagExtExampleLeafModuleToString(i_etDiagExt := iq_stException.udiDiagExt);
TPL.FC_SetException(	i_xExceptionActive	:= TRUE,
						iq_stException		:= iq_stException,
						iq_stExceptionList	:= iq_stExceptionList,
						iq_stLogDataList	:= iq_stLogDataList,
						q_etDiag 			=> etDiagBuffer,
						q_etDiagExt 		=> etDiagExtBufferTPL,
						q_sMsg 				=> sDiagMsgBuffer);

IF (etDiagBuffer <> GD.ET_Diag.Ok) THEN
	(* if exception could not be reported, show exception on outputs *)
	xNotAbleToSetException := TRUE;
	iq_stStandardModuleItf.q_etDiag := iq_stException.etDiag;
	iq_stStandardModuleItf.q_udiDiagExt := iq_stException.udiDiagExt;
	iq_stStandardModuleItf.q_sDiagExt := iq_stException.sDiagExt;
	iq_stStandardModuleItf.q_sMsg := iq_stException.sMsg;
END_IF

stLocalReaction.axReaction[TPL.ET_Reaction.MainsContactorOff] := stLocalReaction.axReaction[TPL.ET_Reaction.MainsContactorOff] OR iq_stException.stReaction.axReaction[TPL.ET_Reaction.MainsContactorOff];
stLocalReaction.axReaction[TPL.ET_Reaction.AsyncStop] := stLocalReaction.axReaction[TPL.ET_Reaction.AsyncStop] OR iq_stException.stReaction.axReaction[TPL.ET_Reaction.AsyncStop];
stLocalReaction.axReaction[TPL.ET_Reaction.SyncStopEH] := stLocalReaction.axReaction[TPL.ET_Reaction.SyncStopEH] OR iq_stException.stReaction.axReaction[TPL.ET_Reaction.SyncStopEH];
stLocalReaction.axReaction[TPL.ET_Reaction.SyncStopEL] := stLocalReaction.axReaction[TPL.ET_Reaction.SyncStopEL] OR iq_stException.stReaction.axReaction[TPL.ET_Reaction.SyncStopEL];
(* special handling for StopEndOfCycle. Wait till reaction feedback from machine. User can transform this reaction and make own reaction.
stLocalReaction.axReaction[TPL.ET_Reaction.StopEndOfCycle] := stLocalReaction.axReaction[TPL.ET_Reaction.StopEndOfCycle] OR iq_stException.stReaction.axReaction[TPL.ET_Reaction.StopEndOfCycle];
*)

stModuleReaction.axReaction[TPL.ET_Reaction.MainsContactorOff] := stLocalReaction.axReaction[TPL.ET_Reaction.MainsContactorOff] OR stModuleReaction.axReaction[TPL.ET_Reaction.MainsContactorOff];
stModuleReaction.axReaction[TPL.ET_Reaction.AsyncStop] := stLocalReaction.axReaction[TPL.ET_Reaction.AsyncStop] OR stModuleReaction.axReaction[TPL.ET_Reaction.AsyncStop];
stModuleReaction.axReaction[TPL.ET_Reaction.SyncStopEH] := stLocalReaction.axReaction[TPL.ET_Reaction.SyncStopEH] OR stModuleReaction.axReaction[TPL.ET_Reaction.SyncStopEH];
stModuleReaction.axReaction[TPL.ET_Reaction.SyncStopEL] := stLocalReaction.axReaction[TPL.ET_Reaction.SyncStopEL] OR stModuleReaction.axReaction[TPL.ET_Reaction.SyncStopEL];
(* special handling for StopEndOfCycle. Wait till reaction feedback from machine. User can transform this reaction and make own reaction.
stModuleReaction.axReaction[TPL.ET_Reaction.StopEndOfCycle] := stLocalReaction.axReaction[TPL.ET_Reaction.StopEndOfCycle] OR stModuleReaction.axReaction[TPL.ET_Reaction.StopEndOfCycle];
*)

(* ---- SetInterfaces.meth.st ---- *)
METHOD SetInterfaces
VAR_INPUT
END_VAR

IF NOT SYSTEMINTERFACE.FC_IsStLogicalAddressValid(i_stLogAddr := iq_stExampleLeafModuleItf.i_ifDrive.stLogicalAddress) THEN
	stExceptionModuleReaction1.etDiag		:= GD.ET_Diag.InputParameterInvalid;
	stExceptionModuleReaction1.udiDiagExt	:= ET_DiagExtExampleLeafModule.DriveInvalid;
	stExceptionModuleReaction1.sMsg			:= 'i_ifDrive - Invalid logical address.';

	ReportException(iq_stException := stExceptionModuleReaction1);
END_IF

xSuccess := __QUERYINTERFACE(iq_stExampleLeafModuleItf.i_ifDrive, ifRefActualValuesPosition);
IF NOT xSuccess OR ifRefActualValuesPosition = 0 THEN
	stExceptionModuleReaction1.etDiag		:= GD.ET_Diag.InputParameterInvalid;
	stExceptionModuleReaction1.udiDiagExt	:= ET_DiagExtExampleLeafModule.DriveInvalid;
	stExceptionModuleReaction1.sMsg			:= 'i_ifDrive : IF_RefActualValues not implemented.';

	ReportException(iq_stException := stExceptionModuleReaction1);
END_IF

(* ---- SetOutputs.meth.st ---- *)
METHOD SetOutputs
VAR_INPUT
END_VAR

IF xNotAbleToSetException THEN
	; (* Do nothing. Diag outputs show not reportable exception *)
	iq_stStandardModuleItf.q_xReady := FALSE;
ELSIF stModuleReaction.axReaction[TPL.ET_Reaction.AsyncStop] THEN
	iq_stStandardModuleItf.q_etDiag := GD.ET_Diag.ExecutionAborted;
	iq_stStandardModuleItf.q_udiDiagExt := ET_DiagExtExampleLeafModule.AsyncStop;
	iq_stStandardModuleItf.q_sDiagExt := 'AsyncStop';
	iq_stStandardModuleItf.q_sMsg := '';

	iq_stStandardModuleItf.q_xReady := FALSE;
ELSIF stModuleReaction.axReaction[TPL.ET_Reaction.SyncStopEL] THEN
	iq_stStandardModuleItf.q_etDiag := GD.ET_Diag.ExecutionAborted;
	iq_stStandardModuleItf.q_udiDiagExt := ET_DiagExtExampleLeafModule.SyncStopEL;
	iq_stStandardModuleItf.q_sDiagExt := 'SyncStopEL';
	iq_stStandardModuleItf.q_sMsg := '';

	iq_stStandardModuleItf.q_xReady := FALSE;
ELSIF stModuleReaction.axReaction[TPL.ET_Reaction.SyncStopEH] THEN
	iq_stStandardModuleItf.q_etDiag := GD.ET_Diag.ExecutionAborted;
	iq_stStandardModuleItf.q_udiDiagExt := ET_DiagExtExampleLeafModule.SyncStopEH;
	iq_stStandardModuleItf.q_sDiagExt := 'SyncStopEH';
	iq_stStandardModuleItf.q_sMsg := '';

	iq_stStandardModuleItf.q_xReady := FALSE;
ELSIF stModuleReaction.axReaction[TPL.ET_Reaction.StopEndOfCycle] THEN
	iq_stStandardModuleItf.q_etDiag := GD.ET_Diag.ExecutionAborted;
	iq_stStandardModuleItf.q_udiDiagExt := ET_DiagExtExampleLeafModule.StopEndOfCycle;
	iq_stStandardModuleItf.q_sDiagExt := 'StopEndOfCycle';
	iq_stStandardModuleItf.q_sMsg := '';

	iq_stStandardModuleItf.q_xReady := FALSE;
ELSE
	IF (iq_stExampleLeafModuleItf.q_etState <> ET_ExampleLeafModuleState.Disabled) AND
	   (iq_stExampleLeafModuleItf.q_etState <> ET_ExampleLeafModuleState.Initializing) THEN

		iq_stStandardModuleItf.q_xReady := TRUE;
	ELSE
		iq_stStandardModuleItf.q_xReady := FALSE;
	END_IF

	iq_stStandardModuleItf.q_etDiag := GD.ET_Diag.Ok;
	CASE iq_stExampleLeafModuleItf.q_etState OF
		ET_ExampleLeafModuleState.NoOp:
			iq_stStandardModuleItf.q_udiDiagExt := ET_DiagExtExampleLeafModule.NoOp;
		ET_ExampleLeafModuleState.Disabled:
			iq_stStandardModuleItf.q_udiDiagExt := ET_DiagExtExampleLeafModule.Disabled;
		ET_ExampleLeafModuleState.Initializing:
			iq_stStandardModuleItf.q_udiDiagExt := ET_DiagExtExampleLeafModule.Initializing;
		ET_ExampleLeafModuleState.HomingWaitForStart:
			iq_stStandardModuleItf.q_udiDiagExt := ET_DiagExtExampleLeafModule.HomingWaitForStart;
		ET_ExampleLeafModuleState.HomingExecuting:
			iq_stStandardModuleItf.q_udiDiagExt := ET_DiagExtExampleLeafModule.HomingExecuting;
		ET_ExampleLeafModuleState.HomingDone:
			iq_stStandardModuleItf.q_udiDiagExt := ET_DiagExtExampleLeafModule.HomingDone;
		ET_ExampleLeafModuleState.AutoWaitForStart:
			iq_stStandardModuleItf.q_udiDiagExt := ET_DiagExtExampleLeafModule.AutoWaitForStart;
		ET_ExampleLeafModuleState.AutoRunning:
			iq_stStandardModuleItf.q_udiDiagExt := ET_DiagExtExampleLeafModule.AutoRunning;
	END_CASE
	iq_stStandardModuleItf.q_sDiagExt := FC_EtDiagExtExampleLeafModuleToString(i_etDiagExt := iq_stStandardModuleItf.q_udiDiagExt);
	iq_stStandardModuleItf.q_sMsg := '';
END_IF

IF fbLoggerPoint.etLogLevel >= APL.ET_LogLevel.StatusMessage THEN
	IF (iq_stExampleLeafModuleItf.q_etState <> etStateOld) THEN
		fbLoggerPoint.AddLogEntry(	i_etLogLevel	:= APL.ET_LogLevel.StatusMessage,
									i_etDiag		:= GD.ET_Diag.Ok,
									i_udiDiagExt	:= ET_DiagExtExampleLeafModule.Ok,
									i_sMessage		:= Standard.CONCAT('State changed to: ', FC_EtExampleLeafModuleStateToString(i_etState := iq_stExampleLeafModuleItf.q_etState)),
									q_etDiag		:= ,
									q_etDiagExt		:= );
	END_IF
	etStateOld := iq_stExampleLeafModuleItf.q_etState;
END_IF

(* ---- SignalSuccessfulExecution.act.st ---- *)
__METADATA__
{
  "v3Meta": {
    "objectGuid": "dc4ccc91-1945-4d06-b781-6fa81c2cc76d",
    "objectTypeGuid": "8ac092e5-3128-4e26-9e7e-11016c6684f2",
    "embeddedObjectTypeGuids": [
      "3b83b776-fb25-43b8-99f2-3c507c9143fc"
    ],
    "properties": {},
    "subObjects": {}
  }
}

IF fbLoggerPoint.etLogLevel >= APL.ET_LogLevel.StatusMessage THEN
	fbLoggerPoint.AddLogEntry(	i_etLogLevel	:= APL.ET_LogLevel.StatusMessage,
								i_etDiag		:= GD.ET_Diag.Ok,
								i_udiDiagExt	:= ET_DiagExtExampleLeafModule.Ok,
								i_sMessage		:= Standard.CONCAT(Standard.CONCAT(Standard.CONCAT('Command done: ', FC_etExampleLeafModuleCmdToString(i_diCmd := iq_stStandardModuleItf.iq_diCmd)),' number: '),DINT_TO_STRING(iq_stStandardModuleItf.iq_diCmd)),
								q_etDiag		:= ,
								q_etDiagExt		:= );
END_IF

iq_stStandardModuleItf.q_xCMDActive := FALSE;
iq_stStandardModuleItf.q_xCMDDone := TRUE;
IF(iq_stStandardModuleItf.iq_diCMD = iq_stStandardModuleItf.q_diCMDActive) THEN
	iq_stStandardModuleItf.iq_diCMD := 0;
(* ELSE don't touch iq_diCMD *)
END_IF

(* ---- SignalUnSuccessfulExecution.act.st ---- *)
__METADATA__
{
  "v3Meta": {
    "objectGuid": "95367f4a-7e78-42be-9529-bfb51b8046a9",
    "objectTypeGuid": "8ac092e5-3128-4e26-9e7e-11016c6684f2",
    "embeddedObjectTypeGuids": [
      "3b83b776-fb25-43b8-99f2-3c507c9143fc"
    ],
    "properties": {},
    "subObjects": {}
  }
}

IF fbLoggerPoint.etLogLevel >= APL.ET_LogLevel.StatusMessage THEN
	fbLoggerPoint.AddLogEntry(	i_etLogLevel	:= APL.ET_LogLevel.StatusMessage,
								i_etDiag		:= GD.ET_Diag.Ok,
								i_udiDiagExt	:= ET_DiagExtExampleLeafModule.Ok,
								i_sMessage		:= Standard.CONCAT(Standard.CONCAT(Standard.CONCAT('Command failed: ', FC_etExampleLeafModuleCmdToString(i_diCmd := iq_stStandardModuleItf.iq_diCmd)),' number: '),DINT_TO_STRING(iq_stStandardModuleItf.iq_diCmd)),
								q_etDiag		:= ,
								q_etDiagExt		:= );
END_IF

iq_stStandardModuleItf.q_xCMDActive := FALSE;
iq_stStandardModuleItf.q_xCMDDone := FALSE;
IF(iq_stStandardModuleItf.iq_diCMD = iq_stStandardModuleItf.q_diCMDActive) THEN
	iq_stStandardModuleItf.iq_diCMD := - iq_stStandardModuleItf.iq_diCMD;
(* ELSE don't touch iq_diCMD *)
END_IF
